Universal Robots URScript: MainCall.script

def MainCall():
  # Global parameters:
  global speed_ms    = 0.250
  global speed_rads  = 0.750
  global accel_mss   = 1.200
  global accel_radss = 1.200
  global blend_radius_m = 0.000

  #--------------------------
  # Add any default subprograms here
  # For example, to drive a gripper as a program call:
  # def Gripper_Open():
  #   ...
  # end
  #
  # Example to drive a spray gun:
  def SprayOn(value):
    # use the value as an output:
    DO_SPRAY = 5
    if value == 0:
      set_standard_digital_out(DO_SPRAY, False)
    else:
      set_standard_digital_out(DO_SPRAY, True)
    end
  end

  # Example to synchronize 2
  def Synchronize():
    # Use the following digital output to signal the state of the robot:
    DO_SYNC = 1

    # Use the following digital input to get the state of another robot:
    DI_SYNC = 1

    if (get_standard_digital_out(DO_SYNC) == get_standard_digital_in(DI_SYNC)):
      set_standard_digital_out(DO_SYNC, not (get_standard_digital_out(DI_SYNC)))
      sleep(0.1)
      thread Thread_wait_1():
        while (True):
          sleep(0.01)
        end
      end
      if (get_standard_digital_out(DO_SYNC) != get_standard_digital_in(DI_SYNC)):
        global thread_handler_1=run Thread_wait_1()
        while (get_standard_digital_out(DO_SYNC) != get_standard_digital_in(DI_SYNC)):
          sync()
        end
        kill thread_handler_1
      end
    else:
      if (get_standard_digital_out(DO_SYNC) != get_standard_digital_in(DI_SYNC)):
        set_standard_digital_out(DO_SYNC, not (get_standard_digital_out(DO_SYNC)))
      end
    end
  end

  #
  # Example to move an external axis
  def MoveAxis(value):
    # use the value as an output:
    DO_AXIS_1 = 1
    DI_AXIS_1 = 1
    if value <= 0:
      set_standard_digital_out(DO_AXIS_1, False)

      # Wait for digital input to change state
      #while (get_standard_digital_in(DI_AXIS_1) != False):
      #  sync()
      #end
    else:
      set_standard_digital_out(DO_AXIS_1, True)

      # Wait for digital input to change state
      #while (get_standard_digital_in(DI_AXIS_1) != True):
      #  sync()
      #end
    end
  end
  #--------------------------

  # Subprogram SubProg2
  def SubProg2():
    movej([0.349066, -0.174533, 0.349066, 0.000000, 0.523599, 0.000000],1.20000,0.75000,0,0.0000)
  end


  # Main program:
  # Program generated by RoboDK v6.0.7 for ABB IRB 120-3/0.6 on XX/XX/XXXX 18:00:00
  # Using nominal kinematics.
  # Using Ref. Frame S: p[1.234570, -0.098765, 0.050500, 0.000000, 0.000000, 0.523599]
  # set_reference(p[1.234570, -0.098765, 0.050500, 0.000000, 0.000000, 0.523599])
  movej([0.000000, -0.174533, 0.349066, 0.000000, 0.523599, 0.000000],1.20000,0.75000,0,0.0000)
  SubProg2()
  NotAProgram()
  # End of main program
end

MainCall()
